Fanuc KAREL source: KT00196.KL

PROGRAM KT00196
%NOLOCKGROUP
VAR
  B1: BOOLEAN
  I2: INTEGER
  OUT: INTEGER
BEGIN
  B1 = TRUE
    I2 = 3
  OUT = B1 AND I2
END KT00196
